TYPE ET_Gr05Manual :
(
	ET_Gr05Manual_eWaitExecute := 0,
	ET_Gr05Manual_eDone := 197,
	ET_Gr05Manual_eError := 198,
	ET_Gr05Manual_eNoExecute := 199
);
END_TYPE

(* stored: Version 1.1.0.1, ProductVersion 3.1.4024.15
   DUT ET_Gr05Manual: Id {1371c67d-cf85-4d0d-8548-2b81b7d6da69} *)
